Fanuc KAREL source: kd00012.KL

PROGRAM KD00012
%STACKSIZE=65535
%PRIORITY=65535
%NOLOCKGROUP
VAR
I : INTEGER
J : INTEGER
B : BOOLEAN
R : REAL
S : STRING[80]
BEGIN
-- UNRESOLVED_PC line 10 opcodes [9D 9D 1A] marker_code=0
END KD00012
